TYPE "FRK_TestResult"
VERSION : 0.1
   STRUCT
      Checks : Int;
      Failures : Int;
      FirstFailure : Int;
      Failed : Array[1..512] of Bool;
      ProtocolError : Bool;
   END_STRUCT;

END_TYPE

